(* IEC 61131-3 sources: BODAS-HelloWorld/st/bodas_rc18_12_40/plc_logic/application, 2 files *)

(* ---- globalvariables-GlobalVariables.st ---- *)
(* --- Interface --- *)
VAR_GLOBAL
	PrmAsw_gstruc             : struc_para;
	anValue_perc_gu8          : USINT;
	swtStatus_gu8             : USINT;
	can1RxDataboxCbkCntr_gu32 : UDINT;
END_VAR
VAR_GLOBAL CONSTANT
	PrmAsw_cgstruc : struc_para := (fctPmp_s16       := 0,
		                            listCtrlVlv_enu  := 1,
		                            nrCogs_s16       := 33,
		                            iSpSafout1_u16   := 500,
		                            iSpSafout2_u16   := 500,
		                            eff_perc_au16    := [10, 50, 90],
		                            nEngSpd_rpm_au16 := [500, 2000, 3500],
		                            PrmDbg_struc     := (flgXcpOn_b := FALSE, flgStoreDataToNvm_b := FALSE));
	ErrMemMgr_nrDfesEntries_DU8 : USINT := 32; (* Maximum number OF errors in DFES *)
	ErrMemMgr_stNoEntryAvl_DU8  : USINT := 255;
	(* bit masks for error states *)
	ErrMemMgr_BitMaskErrDeactvNotSave_DU8 : BYTE := 16#01; (* mask TO fetch Deactive errors which are NOT saved yet *)
	ErrMemMgr_BitMaskErrPrevActv_DU8      : BYTE := 16#10; (* mask TO fetch previously active errors *)
	ErrMemMgr_BitMaskErrActv_DU8          : BYTE := 16#03; (* mask TO fetch active errors *)
	ErrMemMgr_BitMaskErrDeactvSaved_DU8   : BYTE := 16#04; (* mask TO fetch saved deactive errors *)
	ErrMemMgr_BitMaskErrSts_DU8           : BYTE := 16#FF; (* default mask *)
	ErrMemMgr_nrMaxErrEntry_DU8           : BYTE := 27;    (* Max. number of entries, before deleting starts *)
END_VAR

(* ---- main_task_prg-MAIN_TASK_PRG.st ---- *)
(* --- Interface --- *)
(*********************************************************************************************************************
 *    __   __   ___  ___           __   __        __   __  ___
 *   /_ / /  / /__  /    /__/     /_ / /_   |_ / /_ / /  /  /  /__/
 *  /__/ /__/ __ / /__  /  /     /  | /__  /  | /  | /__/  /  /  /
 *
 * Project: Hello World for ml290.rts
 *
 * Program: Main_Task_PRG
 *
 * Description:
 * Main loop of application
 *
 * (c) Copyright by BOSCH REXROTH AG, all rights reserved
 *
 *********************************************************************************************************************)
PROGRAM MAIN_TASK_PRG
VAR
	(******************************************************************************)
	(*************************** _Init ********************************************)
	(******************************************************************************)
	(******************************************************************************)
	(*************************** _Starlock ****************************************)
	(******************************************************************************)
	StartRelease_st_b : BOOL; (*State of the startlock: 1 = the program runs*)
	(******************************************************************************)
	(*************************** _Run *********************************************)
	(******************************************************************************)
	(******************************************************************************)
	(*************************** _PostRun *****************************************)
	(******************************************************************************)
	PostRun_st_b         : BOOL; (*State of the postrun: 1 = the post runs*)
	CallPostRunNr_no_u16 : UINT;
	States_s             : bds_sys_states_ts;
	(******************************************************************************)
	(*************************** _Errors ******************************************)
	(******************************************************************************)
	(******************************************************************************)
	(*************************** _CAN *********************************************)
	(******************************************************************************)
	(******************************************************************************)
	(*************************** General ******************************************)
	(******************************************************************************)
	st_Startlock_b    : BOOL;
	MainTaskState_enu : enu_MainTaskState :=
		enu_MainTaskState.MT_INIT; (* variable indicating the mode of the main task callback function (MT_INIT, MT_CYCLE) *)
END_VAR
VAR CONSTANT
	DELAY_STANDARD       : INT  := 2000; (* debouncing time 2000[ms]*)
	TaskCycleTime_ms_u16 : UINT := 10;   (* Task Cycle Time *)
END_VAR

(* --- Implementation --- *)
CASE MainTaskState_enu OF
enu_MainTaskState.MT_INIT:
	(* Initialization state - only once *)
	INIT();
	StartRelease_st_b := FALSE;
	MainTaskState_enu := enu_MainTaskState.MT_CYCLE;
	ELSE (* -> MT_CYCLE and default state *)
		(* Cyclic state *)
		(* Read inputs *)
		INPUTS();

		IF (StartRelease_st_b) THEN
			IF (PostRun_st_b) THEN
				(* Postrun *)
				POSTRUN();
			ELSE
				(* Normal operational mode *)
				//_RUN();
			END_IF
		ELSE
			(* Wait for start release *)
			STARTLOCK();
		END_IF

		(* Set CAN outputs *)
		CAN_OUT();
		(* Error management *)
		ERRORS();
		(* Set outputs *)
		OUTPUTS();
		(* Reads the parameter from EEPROM *)
		READ_PARAMETERS();
END_CASE
